INTERFACE I_PoseSource

METHOD Reset
VAR_INPUT
	pose : Pose2D;
END_VAR
END_METHOD

PROPERTY Pose : Pose2D
GET
END_GET
END_PROPERTY

END_INTERFACE

(* stored: Version 1.1.0.1, ProductVersion 3.1.4026.12
   Itf I_PoseSource: Id {fb70a82b-2831-5665-93f3-2881a854f361}
   Method Reset: Id {68376bf4-0338-5126-87bc-d465cce5f941}
   Property Pose: Id {88aa799a-c339-5238-aa7c-67fef27207b4}
   Get Get: Id {f2b66024-e9ae-5d09-ba32-37c6a461ad2d} *)
